PROGRAM PMPS_Arbiter
VAR

    fbSetPE	:	PE_Ranges;

    fbBPRequestor : FB_BPRequestor; // Updates global PMPS RequestedBeamParams
    {attribute 'pytmc' := '
    pv: @(PREFIX)PhotonEnergyWatcher
    '}
    fbPhotonEnergyWatcher	:	FB_PhotonEnergyWatcher;

    {attribute 'pytmc' := '
    pv: @(PREFIX)CuRateOutputs
    '}
    fbCuInterface	:	FB_CTLS_Outputs;


    {attribute 'pytmc' := '
    pv: @(PREFIX)BeamParamCntl
    '}
    fbBPControl : FB_BPControlDevice(nID:=16#FFFF);

    (* Subsystem requests use this FB and a pragma link to pass their requests to the arbiter.
    The fb is called on each cycle and updates the arbiter with the current BP set requested
    from the subsystem PLC.*)
    //<TODO> make this so it does input and output to the IF
    (*{attribute 'pytmc' := '
    pv: @(PREFIX):PLC1
    '}*)
    {attribute 'TcLinkTo' := '.i_RequestedBP:=TIIB[plc-kfe-motion]^IO Inputs^RequestedBP;
                                .o_CurrentBP:=TIIB[plc-kfe-motion]^IO Outputs^CurrentBP;
                                .i_Connected:=TIIB[plc-kfe-motion]^SYNC Inputs^External device not connected;
                                .i_WcState:=TIIB[plc-kfe-motion]^WcState^WcStateIn;
                                .i_TxPDOState:=TIIB[plc-kfe-motion]^SYNC Inputs^TxPDO state;
                                '}
    plc_kfe_motion_PMPS_IO : FB_ArbiterToSubSys_IO := (RequestingSystemID := 16#FF0F);




    {attribute 'TcLinkTo' := '.i_RequestedBP:=TIIB[plc-kfe-vac]^IO Inputs^RequestedBP;
                                .o_CurrentBP:=TIIB[plc-kfe-vac]^IO Outputs^CurrentBP;
                                .i_Connected:=TIIB[plc-kfe-vac]^SYNC Inputs^External device not connected;
                                .i_WcState:=TIIB[plc-kfe-vac]^WcState^WcStateIn;
                                .i_TxPDOState:=TIIB[plc-kfe-vac]^SYNC Inputs^TxPDO state;
                                '}
    plc_kfe_vac_PMPS_IO : FB_ArbiterToSubSys_IO := (RequestingSystemID := 16#FF11);

    {attribute 'TcLinkTo' := '.i_RequestedBP:=TIIB[plc-kfe-gatt]^IO Inputs^RequestedBP;
                                .o_CurrentBP:=TIIB[plc-kfe-gatt]^IO Outputs^CurrentBP;
                                .i_Connected:=TIIB[plc-kfe-gatt]^SYNC Inputs^External device not connected;
                                .i_WcState:=TIIB[plc-kfe-gatt]^WcState^WcStateIn;
                                .i_TxPDOState:=TIIB[plc-kfe-gatt]^SYNC Inputs^TxPDO state;
                                '}
    plc_kfe_gatt_PMPS_IO : FB_ArbiterToSubSys_IO := (RequestingSystemID := 16#FF12);

    {attribute 'TcLinkTo' := '.i_RequestedBP:=TIIB[plc-kfe-gmd-vac-01]^IO Inputs^RequestedBP;
                                .o_CurrentBP:=TIIB[plc-kfe-gmd-vac-01]^IO Outputs^CurrentBP;
                                .i_Connected:=TIIB[plc-kfe-gmd-vac-01]^SYNC Inputs^External device not connected;
                                .i_WcState:=TIIB[plc-kfe-gmd-vac-01]^WcState^WcStateIn;
                                .i_TxPDOState:=TIIB[plc-kfe-gmd-vac-01]^SYNC Inputs^TxPDO state;
                                '}
    plc_kfe_gmd_PMPS_IO : FB_ArbiterToSubSys_IO := (RequestingSystemID := 16#FF13);

    {attribute 'TcLinkTo' := '.i_RequestedBP:=TIIB[plc-kfe-xgmd-vac-01]^IO Inputs^RequestedBP;
                                .o_CurrentBP:=TIIB[plc-kfe-xgmd-vac-01]^IO Outputs^CurrentBP;
                                .i_Connected:=TIIB[plc-kfe-xgmd-vac-01]^SYNC Inputs^External device not connected;
                                .i_WcState:=TIIB[plc-kfe-xgmd-vac-01]^WcState^WcStateIn;
                                .i_TxPDOState:=TIIB[plc-kfe-xgmd-vac-01]^SYNC Inputs^TxPDO state;
                                '}
    plc_kfe_xgmd_PMPS_IO : FB_ArbiterToSubSys_IO := (RequestingSystemID := 16#FF14);



//////////////////////////////////////////////
// TMO PLCs
/////////////////////////////////////////////

    {attribute 'TcLinkTo' := '.i_RequestedBP:=TIIB[plc-tmo-mot]^IO Inputs^RequestedBP;
                                .o_CurrentBP:=TIIB[plc-tmo-mot]^IO Outputs^CurrentBP;
                                .i_Connected:=TIIB[plc-tmo-mot]^SYNC Inputs^External device not connected;
                                .i_WcState:=TIIB[plc-tmo-mot]^WcState^WcStateIn;
                                .i_TxPDOState:=TIIB[plc-tmo-mot]^SYNC Inputs^TxPDO state;
                                '}
    plc_tmo_motion_PMPS_IO : FB_ArbiterToSubSys_IO := (RequestingSystemID := 16#F100);

    {attribute 'TcLinkTo' := '.i_RequestedBP:=TIIB[plc-tmo-optics]^IO Inputs^RequestedBP;
                                .o_CurrentBP:=TIIB[plc-tmo-optics]^IO Outputs^CurrentBP;
                                .i_Connected:=TIIB[plc-tmo-optics]^SYNC Inputs^External device not connected;
                                .i_WcState:=TIIB[plc-tmo-optics]^WcState^WcStateIn;
                                .i_TxPDOState:=TIIB[plc-tmo-optics]^SYNC Inputs^TxPDO state;
                                '}
    plc_tmo_optics_PMPS_IO : FB_ArbiterToSubSys_IO := (RequestingSystemID := 16#F101);

    {attribute 'TcLinkTo' := '.i_RequestedBP:=TIIB[plc-tmo-vac]^IO Inputs^RequestedBP;
                                .o_CurrentBP:=TIIB[plc-tmo-vac]^IO Outputs^CurrentBP;
                                .i_Connected:=TIIB[plc-tmo-vac]^SYNC Inputs^External device not connected;
                                .i_WcState:=TIIB[plc-tmo-vac]^WcState^WcStateIn;
                                .i_TxPDOState:=TIIB[plc-tmo-vac]^SYNC Inputs^TxPDO state;
                                '}
    plc_tmo_vacuum_PMPS_IO : FB_ArbiterToSubSys_IO := (RequestingSystemID := 16#F102);

    count : CTU;
//////////////////////////////////////////////
// RIX PLCs
/////////////////////////////////////////////
    {attribute 'TcLinkTo' := '.i_RequestedBP:=TIIB[plc-rix-vac]^IO Inputs^RequestedBP;
                                .o_CurrentBP:=TIIB[plc-rix-vac]^IO Outputs^CurrentBP;
                                .i_Connected:=TIIB[plc-rix-vac]^SYNC Inputs^External device not connected;
                                .i_WcState:=TIIB[plc-rix-vac]^WcState^WcStateIn;
                                .i_TxPDOState:=TIIB[plc-rix-vac]^SYNC Inputs^TxPDO state;
                                '}
    plc_rix_vac_PMPS_IO : FB_ArbiterToSubSys_IO := (RequestingSystemID := 16#F200);

    {attribute 'TcLinkTo' := '.i_RequestedBP:=TIIB[plc-rix-optics]^IO Inputs^RequestedBP;
                                .o_CurrentBP:=TIIB[plc-rix-optics]^IO Outputs^CurrentBP;
                                .i_Connected:=TIIB[plc-rix-optics]^SYNC Inputs^External device not connected;
                                .i_WcState:=TIIB[plc-rix-optics]^WcState^WcStateIn;
                                .i_TxPDOState:=TIIB[plc-rix-optics]^SYNC Inputs^TxPDO state;
                                '}
    plc_rix_optics_PMPS_IO : FB_ArbiterToSubSys_IO := (RequestingSystemID := 16#F201);

    {attribute 'TcLinkTo' := '.i_RequestedBP:=TIIB[plc-rix-mot]^IO Inputs^RequestedBP;
                                .o_CurrentBP:=TIIB[plc-rix-mot]^IO Outputs^CurrentBP;
                                .i_Connected:=TIIB[plc-rix-mot]^SYNC Inputs^External device not connected;
                                .i_WcState:=TIIB[plc-rix-mot]^WcState^WcStateIn;
                                .i_TxPDOState:=TIIB[plc-rix-mot]^SYNC Inputs^TxPDO state;
                                '}
    plc_rix_mot_PMPS_IO : FB_ArbiterToSubSys_IO := (RequestingSystemID := 16#F202);

    {attribute 'TcLinkTo' := '.i_RequestedBP:=TIIB[plc-crix-mot]^IO Inputs^RequestedBP;
                                .o_CurrentBP:=TIIB[plc-crix-mot]^IO Outputs^CurrentBP;
                                .i_Connected:=TIIB[plc-crix-mot]^SYNC Inputs^External device not connected;
                                .i_WcState:=TIIB[plc-crix-mot]^WcState^WcStateIn;
                                .i_TxPDOState:=TIIB[plc-crix-mot]^SYNC Inputs^TxPDO state;
                                '}
    plc_crix_mot_PMPS_IO : FB_ArbiterToSubSys_IO := (RequestingSystemID := 16#F203);

{attribute 'TcLinkTo' := '.i_RequestedBP:=TIIB[plc-crix-vac]^IO Inputs^RequestedBP;
                                .o_CurrentBP:=TIIB[plc-crix-vac]^IO Outputs^CurrentBP;
                                .i_Connected:=TIIB[plc-crix-vac]^SYNC Inputs^External device not connected;
                                .i_WcState:=TIIB[plc-crix-vac]^WcState^WcStateIn;
                                .i_TxPDOState:=TIIB[plc-crix-vac]^SYNC Inputs^TxPDO state;
                                '}
    plc_crix_vac_PMPS_IO : FB_ArbiterToSubSys_IO := (RequestingSystemID := 16#F205);

    {attribute 'TcLinkTo' := '.i_RequestedBP:=TIIB[plc-qrix-mot]^IO Inputs^RequestedBP;
                                .o_CurrentBP:=TIIB[plc-qrix-mot]^IO Outputs^CurrentBP;
                                .i_Connected:=TIIB[plc-qrix-mot]^SYNC Inputs^External device not connected;
                                .i_WcState:=TIIB[plc-qrix-mot]^WcState^WcStateIn;
                                .i_TxPDOState:=TIIB[plc-qrix-mot]^SYNC Inputs^TxPDO state;
                                '}


    plc_qrix_mot_PMPS_IO : FB_ArbiterToSubSys_IO := (RequestingSystemID := 16#F206);

    {attribute 'TcLinkTo' := '.i_RequestedBP:=TIIB[plc-qrix-vac]^IO Inputs^RequestedBP;
                                .o_CurrentBP:=TIIB[plc-qrix-vac]^IO Outputs^CurrentBP;
                                .i_Connected:=TIIB[plc-qrix-vac]^SYNC Inputs^External device not connected;
                                .i_WcState:=TIIB[plc-qrix-vac]^WcState^WcStateIn;
                                .i_TxPDOState:=TIIB[plc-qrix-vac]^SYNC Inputs^TxPDO state;
                                '}
    plc_qrix_vac_PMPS_IO : FB_ArbiterToSubSys_IO := (RequestingSystemID := 16#F204);

//////////////////////////////////////////////
// TXI PLCs
/////////////////////////////////////////////

    {attribute 'TcLinkTo' := '.i_RequestedBP:=TIIB[plc-txi-mot]^IO Inputs^RequestedBP;
                                .o_CurrentBP:=TIIB[plc-txi-mot]^IO Outputs^CurrentBP;
                                .i_Connected:=TIIB[plc-txi-mot]^SYNC Inputs^External device not connected;
                                .i_WcState:=TIIB[plc-txi-mot]^WcState^WcStateIn;
                                .i_TxPDOState:=TIIB[plc-txi-mot]^SYNC Inputs^TxPDO state;
                                '}
    plc_txi_motion_PMPS_IO : FB_ArbiterToSubSys_IO := (RequestingSystemID := 16#F300);

    {attribute 'TcLinkTo' := '.i_RequestedBP:=TIIB[plc-txi-optics]^IO Inputs^RequestedBP;
                                .o_CurrentBP:=TIIB[plc-txi-optics]^IO Outputs^CurrentBP;
                                .i_Connected:=TIIB[plc-txi-optics]^SYNC Inputs^External device not connected;
                                .i_WcState:=TIIB[plc-txi-optics]^WcState^WcStateIn;
                                .i_TxPDOState:=TIIB[plc-txi-optics]^SYNC Inputs^TxPDO state;
                                '}
    plc_txi_optics_PMPS_IO : FB_ArbiterToSubSys_IO := (RequestingSystemID := 16#F301);

    {attribute 'TcLinkTo' := '.i_RequestedBP:=TIIB[plc-txi-vac]^IO Inputs^RequestedBP;
                                .o_CurrentBP:=TIIB[plc-txi-vac]^IO Outputs^CurrentBP;
                                .i_Connected:=TIIB[plc-txi-vac]^SYNC Inputs^External device not connected;
                                .i_WcState:=TIIB[plc-txi-vac]^WcState^WcStateIn;
                                .i_TxPDOState:=TIIB[plc-txi-vac]^SYNC Inputs^TxPDO state;
                                '}
    plc_txi_vacuum_PMPS_IO : FB_ArbiterToSubSys_IO := (RequestingSystemID := 16#F302);

    (*Remove*)
         ar1 : bool;
 ar2 : bool;
 nReqID:UDINT;
 nReqRM:UDINT;
 bRemove:bool;
 rtRemove: R_TRIG;

END_VAR


// Updating arbiter with subsystem requests.

///////////////////////////
// KFE
    plc_kfe_motion_PMPS_IO(Arbiter:=GVL.g_fbArbiter1, fbFFHWO:=GVL.g_FastFaultOutput1, Reset:=GVL.AttemptReset, sName:= 'KFE MOTION');
    plc_kfe_vac_PMPS_IO(Arbiter:=GVL.g_fbArbiter1, fbFFHWO:=GVL.g_FastFaultOutput1, Reset:=GVL.AttemptReset, sName:= 'KFE VACUUM');
    plc_kfe_gatt_PMPS_IO(Arbiter:=GVL.g_fbArbiter1, fbFFHWO:=GVL.g_FastFaultOutput1, Reset:=GVL.AttemptReset, sName:= 'KFE GATT');
///////////////////////////

///////////////////////////
// TMO K4
// TMO-OPTICS Veto	MR1K1_IN
    plc_tmo_optics_PMPS_IO(Arbiter:=GVL.g_fbArbiter1, fbFFHWO:=GVL.g_FastFaultOutput3, Reset:=GVL.AttemptReset, sName:= 'TMO OPTICS');
// TMO-VAC and TMO-MOT OR ST3K4_IN
    plc_tmo_motion_PMPS_IO(Arbiter:=GVL.g_fbArbiter1, fbFFHWO:=GVL.g_FastFaultOutput4, Reset:=GVL.AttemptReset , sName:= 'TMO MOTION');
    plc_tmo_vacuum_PMPS_IO(Arbiter:=GVL.g_fbArbiter1, fbFFHWO:=GVL.g_FastFaultOutput4, Reset:=GVL.AttemptReset, sName:= 'TMO VACUUM');
///////////////////////////
	
//////////////////////////
// RIX
// RIX- OPTICS No Veto / Should be FFO:01 since it is upstream of all Vetos
	plc_rix_optics_PMPS_IO(Arbiter:=GVL.g_fbArbiter1, fbFFHWO:=GVL.g_FastFaultOutput1, Reset:=GVL.AttemptReset, sName:= 'RIX OPTICS');
// RIX-VAC and RIX-MOT MR1K1_OUT
    plc_rix_vac_PMPS_IO(Arbiter:=GVL.g_fbArbiter1, fbFFHWO:=GVL.g_FastFaultOutput5, Reset:=GVL.AttemptReset, sName:= 'RIX VACUUM'); 
    plc_rix_mot_PMPS_IO(Arbiter:=GVL.g_fbArbiter1, fbFFHWO:=GVL.g_FastFaultOutput5, Reset:=GVL.AttemptReset, sName:= 'RIX MOTION');
// QRIX-VAC, CRIX-VAC and CRIX-MOT MR1K1_OUT OR ST1K2_IN
	plc_crix_mot_PMPS_IO(Arbiter:=GVL.g_fbArbiter1, fbFFHWO:=GVL.g_FastFaultOutput6, Reset:=GVL.AttemptReset, sName:= 'CRIX MOTION');
    plc_crix_vac_PMPS_IO(Arbiter:=GVL.g_fbArbiter1, fbFFHWO:=GVL.g_FastFaultOutput6, Reset:=GVL.AttemptReset, sName:= 'CRIX VACUUM');
    plc_qrix_vac_PMPS_IO(Arbiter:=GVL.g_fbArbiter1, fbFFHWO:=GVL.g_FastFaultOutput6, Reset:=GVL.AttemptReset, sName:= 'QRIX VACUUM');
///////////////////////////


///////////////////////////
// TXI K3
// TXI- OPTICS No Veto / Should be FFO:01 since it is upstream of all Vetos
    plc_txi_optics_PMPS_IO(Arbiter:=GVL.g_fbArbiter1, fbFFHWO:=GVL.g_FastFaultOutput1, Reset:=GVL.AttemptReset, sName:= 'TXI OPTICS');
// TXI-VAC and TXI-MOT 	MR1K3_OUT and MR2K3_OUT
    plc_txi_vacuum_PMPS_IO(Arbiter:=GVL.g_fbArbiter1, fbFFHWO:=GVL.g_FastFaultOutput7, Reset:=GVL.AttemptReset, sName:= 'TXI VACUUM');
	plc_txi_motion_PMPS_IO(Arbiter:=GVL.g_fbArbiter1, fbFFHWO:=GVL.g_FastFaultOutput7, Reset:=GVL.AttemptReset , sName:= 'TXI MOTION');
//////////////////////////


///////////////////////////
//Beam Class override
// Dummy device for controling pmps beam parameters
fbBPControl(Arbiter:=g_fbArbiter2);

//Call the program that evaluates the Override and generate the correct Beam Parameter and adds it to arbiter 2
P_Override_Tran_BC();

////////////////////////////
// Beam parameter requestor
//////////////////////////////
fbBPRequestor(Arbiter:=GVL.g_fbArbiter2, q_ReqBP => PMPS_GVL.stRequestedBeamParameters);

//Now lets write the FAKE BP to send to the PLCs
GVL.stCurrentFakeBP := PMPS_GVL.stCurrentBeamParameters;
IF (bApplyJF) THEN
    //What if we are NOT in override mode? Then the Arbitrated1BP should be the current BP, right?
    //Should we always broadcast the requested arbitratedBP
    // yes and no. I think that it should be either the safer or the ArbitratedBP because of a specific use case in RIX OPTICS
    IF (PMPS_GVL.stCurrentBeamParameters.nTran > GVL.stArbiter1BP.nTran) THEN
        GVL.stCurrentFakeBP.nTran:= GVL.stArbiter1BP.nTran;
    END_IF
    IF (PMPS_GVL.stCurrentBeamParameters.nBeamClass > GVL.stArbiter1BP.nBeamClass) THEN
        GVL.stCurrentFakeBP.nBeamClass:= GVL.stArbiter1BP.nBeamClass;
        GVL.stCurrentFakeBP.nBCRange:= GVL.stArbiter1BP.nBCRange;
    END_IF
END_IF


// Request Cu beam rate
fbCuInterface(BP := PMPS_GVL.stRequestedBeamParameters);


// Keep an eye on the photon energy
fbPhotonEnergyWatcher(i_stCurrentBeamParams	:= PMPS_GVL.stCurrentBeamParameters,
                    i_stRequestedBeamParams := PMPS_GVL.stRequestedBeamParameters,
                    io_fbFFHWO:= GVL.g_FastFaultOutput1,
                    i_xReset := GVL.AttemptReset);

//Assert beam class
P_BeamClassAssertion();


//Use Only in very critical cases. Only when you are sure. This might result in damage to devices
(*remove*)
(*Debugging functions*)
ar1:= GVL.g_fbArbiter1.CheckRequestInPool(nReqRM);

rtRemove(CLK:= bRemove);
if (rtRemove.Q) THEN
     GVL.g_fbArbiter1.RemoveRequest(nReqRM);
END_IF

END_PROGRAM

(* stored: Version 1.1.0.1, ProductVersion 3.1.4022.18
   POU PMPS_Arbiter: Id {91ae890b-11cc-4d41-83ec-edc5b802c784}, SpecialFunc None *)
